(* IEC 61131-3 sources: Grupo7_SParcial_Automatizacion_Control/2. openPLC_file/openPLC_V2.1/build, 2 files *)

(* ---- plc.st ---- *)
TYPE
  LOGLEVEL : (CRITICAL, WARNING, INFO, DEBUG) := INFO;
END_TYPE

FUNCTION_BLOCK LOGGER
  VAR_INPUT
    TRIG : BOOL;
    MSG : STRING;
    LEVEL : LOGLEVEL := INFO;
  END_VAR
  VAR
    TRIG0 : BOOL;
  END_VAR

  IF TRIG AND NOT TRIG0 THEN
  {{
   LogMessage(GetFbVar(LEVEL),(char*)GetFbVar(MSG, .body),GetFbVar(MSG, .len));
  }}
  END_IF;
  TRIG0:=TRIG;
END_FUNCTION_BLOCK

FUNCTION_BLOCK python_eval
  VAR_INPUT
    TRIG : BOOL;
    CODE : STRING;
  END_VAR
  VAR_OUTPUT
    ACK : BOOL;
    RESULT : STRING;
  END_VAR
  VAR
    STATE : DWORD;
    BUFFER : STRING;
    PREBUFFER : STRING;
    TRIGM1 : BOOL;
    TRIGGED : BOOL;
  END_VAR

  {extern void __PythonEvalFB(int, PYTHON_EVAL*);__PythonEvalFB(0, data__);}
END_FUNCTION_BLOCK

FUNCTION_BLOCK python_poll
  VAR_INPUT
    TRIG : BOOL;
    CODE : STRING;
  END_VAR
  VAR_OUTPUT
    ACK : BOOL;
    RESULT : STRING;
  END_VAR
  VAR
    STATE : DWORD;
    BUFFER : STRING;
    PREBUFFER : STRING;
    TRIGM1 : BOOL;
    TRIGGED : BOOL;
  END_VAR

  {extern void __PythonEvalFB(int, PYTHON_EVAL*);__PythonEvalFB(1,(PYTHON_EVAL*)(void*)data__);}
END_FUNCTION_BLOCK

FUNCTION_BLOCK python_gear
  VAR_INPUT
    N : UINT;
    TRIG : BOOL;
    CODE : STRING;
  END_VAR
  VAR_OUTPUT
    ACK : BOOL;
    RESULT : STRING;
  END_VAR
  VAR
    py_eval : python_eval;
    COUNTER : UINT;
    _TMP_ADD10_OUT : UINT;
    _TMP_EQ13_OUT : BOOL;
    _TMP_SEL15_OUT : UINT;
    _TMP_AND7_OUT : BOOL;
  END_VAR

  _TMP_ADD10_OUT := ADD(COUNTER, 1);
  _TMP_EQ13_OUT := EQ(N, _TMP_ADD10_OUT);
  _TMP_SEL15_OUT := SEL(_TMP_EQ13_OUT, _TMP_ADD10_OUT, 0);
  COUNTER := _TMP_SEL15_OUT;
  _TMP_AND7_OUT := AND(_TMP_EQ13_OUT, TRIG);
  py_eval(TRIG := _TMP_AND7_OUT, CODE := CODE);
  ACK := py_eval.ACK;
  RESULT := py_eval.RESULT;
END_FUNCTION_BLOCK

PROGRAM exam_openPLC_simu
  VAR
    s1_arrive : BOOL;
    s2_arrive : BOOL;
    s3_bottle_full : BOOL;
    s4_bottle_seal : BOOL;
    start : BOOL;
    bomb : BOOL;
    Ms_down_up : BOOL;
    M1_M2 : BOOL;
  END_VAR
  VAR
    TON0 : TON;
  END_VAR

  IF start THEN
    M1_M2 := TRUE; (*set*)
  END_IF;
  IF s1_arrive THEN
    M1_M2 := FALSE; (*reset*)
  END_IF;
  IF s1_arrive THEN
    bomb := TRUE; (*set*)
  END_IF;
  IF s3_bottle_full THEN
    bomb := FALSE; (*reset*)
  END_IF;
  IF s3_bottle_full THEN
    M1_M2 := TRUE; (*set*)
  END_IF;
  IF s2_arrive THEN
    M1_M2 := FALSE; (*reset*)
  END_IF;
  IF s2_arrive THEN
    Ms_down_up := TRUE; (*set*)
  END_IF;
  TON0(IN := Ms_down_up, PT := T#1000ms);
  IF TON0.Q THEN
    Ms_down_up := FALSE; (*reset*)
  END_IF;
  IF s4_bottle_seal THEN
    M1_M2 := TRUE; (*set*)
  END_IF;
END_PROGRAM

CONFIGURATION Config0

  RESOURCE Res0 ON PLC
    TASK task0(INTERVAL := T#20ms,PRIORITY := 0);
    PROGRAM instance0 WITH task0 : exam_openPLC_simu;
  END_RESOURCE
END_CONFIGURATION

(* ---- generated_plc.st ---- *)
PROGRAM exam_openPLC_simu
  VAR
    s1_arrive AT %IX0.0 : BOOL;
    s2_arrive AT %IX0.1 : BOOL;
    s3_bottle_full AT %IX0.2 : BOOL;
    s4_bottle_seal AT %IX0.3 : BOOL;
    start AT %IX0.4 : BOOL;
    bomb AT %QX0.0 : BOOL;
    Ms_down_up AT %QX0.1 : BOOL;
    M1_M2 AT %QX0.2 : BOOL;
  END_VAR
  VAR
    TON0 : TON;
  END_VAR

  IF start THEN
    M1_M2 := TRUE; (*set*)
  END_IF;
  IF s1_arrive THEN
    M1_M2 := FALSE; (*reset*)
  END_IF;
  IF s1_arrive THEN
    bomb := TRUE; (*set*)
  END_IF;
  IF s3_bottle_full THEN
    bomb := FALSE; (*reset*)
  END_IF;
  IF s3_bottle_full THEN
    M1_M2 := TRUE; (*set*)
  END_IF;
  IF s2_arrive THEN
    M1_M2 := FALSE; (*reset*)
  END_IF;
  IF s2_arrive THEN
    Ms_down_up := TRUE; (*set*)
  END_IF;
  TON0(IN := Ms_down_up, PT := T#1000ms);
  IF TON0.Q THEN
    Ms_down_up := FALSE; (*reset*)
  END_IF;
  IF s4_bottle_seal THEN
    M1_M2 := TRUE; (*set*)
  END_IF;
END_PROGRAM

CONFIGURATION Config0

  RESOURCE Res0 ON PLC
    TASK task0(INTERVAL := T#20ms,PRIORITY := 0);
    PROGRAM instance0 WITH task0 : exam_openPLC_simu;
  END_RESOURCE
END_CONFIGURATION
